Staubli VAL3: setIOStatus.pgx

public program setIOStatus(num x_nType)
  local num l_nSize
  local string l_selColor
  local string l_sNullColor
  local string l_sbtn
  local string l_sErrColor
  local string l_slabel
  local num l_nValue
  local num l_i
  local num l_nSize1
  local string l_slbl1
  local string l_slbl2
begin
  l_selColor="#33FF33"
  l_sNullColor="#FFFFFF"
  l_sErrColor="#C8C8C8"
  call getSize(l_nSize,l_nSize1)
  //  if l_nSize<16
  //    for l_i = l_nSize to 15
  //      l_sbtn="btn"+toString("",60+l_i)
  //      l_slbl1="lbl"+toString("",20+l_i)
  //      l_slbl2="lbl"+toString("",l_i)
  //      userPageSet("IO",l_sbtn,"style.visibility","hidden")
  //      userPageSet("IO",l_slbl1,"style.visibility","hidden")
  //      userPageSet("IO",l_slbl2,"style.visibility","hidden")
  //    endFor
  //  endIf
  //  if l_nSize1<16
  //    for l_i = l_nSize1 to 15
  //      l_sbtn="lbl"+toString("",40+l_i)
  //      l_slbl1="lbl"+toString("",20+l_i)
  //      l_slbl2="lbl"+toString("",l_i)
  //      userPageSet("IO",l_sbtn,"style.visibility","hidden")
  //      userPageSet("IO",l_slbl1,"style.visibility","hidden")
  //      userPageSet("IO",l_slbl2,"style.visibility","hidden")
  //    endFor
  //  endIf

  switch x_nType
    case 0
      for l_i = 0 to l_nSize-1
        l_sbtn="btn"+toString("",60+l_i)
        //     userPageSet("IO",l_sbtn,"style.visibility","visible")
        if ioStatus(io:dInItem[l_i+nPageIndex*16].dDio)>-1
          l_nValue=dioGet(io:dInItem[l_i+nPageIndex*16].dDio)
          if l_nValue==1
            userPageSet("IO",l_sbtn,"style.backgroundColor",l_selColor)
          else
            userPageSet("IO",l_sbtn,"style.backgroundColor",l_sNullColor)
          endIf
        else
          userPageSet("IO",l_sbtn,"style.backgroundColor",l_sErrColor)
        endIf
      endFor
    break
    case 1
      for l_i = 0 to l_nSize-1
        l_sbtn="btn"+toString("",60+l_i)
        //     userPageSet("IO",l_sbtn,"style.visibility","visible")
        if ioStatus(io:dOutItem[l_i+nPageIndex*16].dDio)>-1
          l_nValue=dioGet(io:dOutItem[l_i+nPageIndex*16].dDio)
          if l_nValue==1
            userPageSet("IO",l_sbtn,"style.backgroundColor",l_selColor)
          else
            userPageSet("IO",l_sbtn,"style.backgroundColor",l_sNullColor)
          endIf
        else
          userPageSet("IO",l_sbtn,"style.backgroundColor",l_sErrColor)
        endIf
      endFor
    break
    case 2
      for l_i = 0 to l_nSize1-1
        l_slabel="lbl"+toString("",40+l_i)
        //       userPageSet("IO",l_slabel,"style.visibility","visible")
        if ioStatus(io:aInItem[l_i+nPageIndex*16].aAio)>-1
          l_nValue=aioGet(io:aInItem[l_i+nPageIndex*16].aAio)
          sValue[l_i]=toString(".2",l_nValue)
        else
          sValue[l_i]="?"
        endIf
      endFor
    break
    case 3
      for l_i = 0 to l_nSize1-1
        l_slabel="lbl"+toString("",40+l_i)
        //      userPageSet("IO",l_slabel,"style.visibility","visible")
        if ioStatus(io:aOutItem[l_i+nPageIndex*16].aAio)>-1
          l_nValue=aioGet(io:aOutItem[l_i+nPageIndex*16].aAio)
          sValue[l_i]=toString(".2",l_nValue)
        else
          sValue[l_i]="?"
        endIf
      endFor
    break

  endSwitch

end
